  # Gripper Configurations depending on the Object Type , add new force and speed in the Defines if necessary
  # create_gripper_config(gripper_offset=struct(prepick=2, pick=0, place=2), force=0, speed=0, validation=0, object=create_object())
  GRIPPER_CONFIG_MAP.append(create_gripper_config(gripper_offset=struct(prepick=2, pick=0, place=2), force=GRIPPER_FORCE.HALF, speed=GRIPPER_SPEED.MEDIUM, validation=GRIPPER_VALIDATION.ON, object=find_object_by_objectname(Objects.ANY_SAMPLE)))
  GRIPPER_CONFIG_MAP.append(create_gripper_config(gripper_offset=struct(prepick=2, pick=0, place=2), force=GRIPPER_FORCE.FULL, speed=GRIPPER_SPEED.MEDIUM, validation=GRIPPER_VALIDATION.ON, object=find_object_by_objectname(Objects.ANY_RACK)))
  GRIPPER_CONFIG_MAP.append(create_gripper_config(gripper_offset=struct(prepick=2, pick=0, place=2), force=GRIPPER_FORCE.HALF, speed=GRIPPER_SPEED.MEDIUM, validation=GRIPPER_VALIDATION.ON, object=find_object_by_objectname(Objects.CC_SAMPLE)))
  GRIPPER_CONFIG_MAP.append(create_gripper_config(gripper_offset=struct(prepick=3, pick=0, place=3), force=GRIPPER_FORCE.HALF, speed=GRIPPER_SPEED.MEDIUM, validation=GRIPPER_VALIDATION.ON, object=find_object_by_objectname(Objects.HEMA_SAMPLE)))
  GRIPPER_CONFIG_MAP.append(create_gripper_config(gripper_offset=struct(prepick=4, pick=0, place=4), force=GRIPPER_FORCE.HALF, speed=GRIPPER_SPEED.MEDIUM, validation=GRIPPER_VALIDATION.OFF, object=find_object_by_objectname(Objects.TARA_SAMPLE)))
  GRIPPER_CONFIG_MAP.append(create_gripper_config(gripper_offset=struct(prepick=2, pick=0, place=2), force=GRIPPER_FORCE.FULL, speed=GRIPPER_SPEED.MEDIUM, validation=GRIPPER_VALIDATION.ON, object=find_object_by_objectname(Objects.CF_RACK)))
  GRIPPER_CONFIG_MAP.append(create_gripper_config(gripper_offset=struct(prepick=2, pick=0, place=2), force=GRIPPER_FORCE.FULL, speed=GRIPPER_SPEED.MEDIUM, validation=GRIPPER_VALIDATION.ON, object=find_object_by_objectname(Objects.COBAS_RACK)))
  GRIPPER_CONFIG_MAP.append(create_gripper_config(gripper_offset=struct(prepick=0, pick=0, place=0), force=GRIPPER_FORCE.HALF, speed=GRIPPER_SPEED.MEDIUM, validation=GRIPPER_VALIDATION.OFF, object=find_object_by_objectname(Objects.NONE)))
  GRIPPER_CONFIG_MAP.append(create_gripper_config(gripper_offset=struct(prepick=0, pick=0, place=0), force=GRIPPER_FORCE.HALF, speed=GRIPPER_SPEED.MEDIUM, validation=GRIPPER_VALIDATION.OFF, object=find_object_by_objectname(Objects.BUTTON)))
  GRIPPER_CONFIG_MAP.append(create_gripper_config(gripper_offset=struct(prepick=5, pick=25, place=5), force=GRIPPER_FORCE.HALF, speed=GRIPPER_SPEED.MEDIUM, validation=GRIPPER_VALIDATION.OFF, object=find_object_by_objectname(Objects.XN550_DRAWER)))
  # create Patterns like Racks or Magazines
  # easy if you define x and y regarding to the base coordinate system  if not you have to deal with transpose and or invert
  # create_pattern(id=0, pattern_width=[0, 0], pattern_size=[0, 0], blocked=[-1, -1], obj_name=0, direction="X", transpose=False, invert=False, description="default")
  # Objectss: NONE=0, CC_SAMPLE=1, CC_RACK=2, COAG_SAMPLE=3, COAG_RACK=4, HEMA_SAMPLE=5, HEMA_RACK=6, INPUT_RACK=7, CENTRIFUGE_RACK=8, ANY_SAMPLE=9, ANY_RACK=10
  # ITEM_MODEL_MAP.append(create_pattern(id=0, pattern_width=[0, 0], pattern_size=[0, 0], blocked=[-1, -1, -1],  direction="X", transpose=False, invert=False, description="default"))
  # ITEM_MODEL_MAP.append(create_pattern(id=1, pattern_width=[0.06, 0], pattern_size=[3, 1],  direction="X", description="Tara"))
  # ITEM_MODEL_MAP.append(create_pattern(id=2, pattern_width=[0.183, 0.082], pattern_size=[10, 5], description="Sarstedt 50 D17 Rack"))
  # ITEM_MODEL_MAP.append(create_pattern(id=3, pattern_width=[0.153, 0.067], pattern_size=[10, 5], description="Sarstedt 50 D13 Rack"))
  # ITEM_MODEL_MAP.append(create_pattern(id=4, pattern_width=[0.06, 0.06], pattern_size=[3, 3], blocked=[5, -1, -1], description="Hettich Centrifuge Rack"))
  # ITEM_MODEL_MAP.append(create_pattern(id=5, pattern_width=[0.093, 0.093], pattern_size=[2, 2],  description="Hettich Centrifuge Rack Magazin"))
  # ITEM_MODEL_MAP.append(create_pattern(id=6, pattern_width=[0.08, 0.05], pattern_size=[5, 2], description="Sysmex XN 550 Rack"))
  # ITEM_MODEL_MAP.append(create_pattern(id=7, pattern_width=[0.175, 0.078], pattern_size=[8, 4], description="URG Rack 40 D17"))
  # ITEM_MODEL_MAP.append(create_pattern(id=8, pattern_width=[0.092, 0], pattern_size=[5, 1], description="Cobas Rack"))
  # ITEM_MODEL_MAP.append(create_pattern(id=9, pattern_width=[0.245, 0.123], pattern_size=[3, 5], blocked=[9,11,12], description="Cobas Rack Magazin"))
  # ITEM_MODEL_MAP.append(create_pattern(id=10, pattern_width=[0.237, 0.095], pattern_size=[11, 5], description="Atellica Rack 5x11"))
  # ITEM_MODEL_MAP.append(create_pattern(id=11, pattern_width=[0.237, 0.095], pattern_size=[2, 2], description="Sensors LM"))
  # ITEM_MODEL_MAP.append(create_pattern(id=12, pattern_width=[0.18, 0], pattern_size=[10, 1], description="Sysmex CS2500 Rack"))
  # ITEM_MODEL_MAP.append(create_pattern(id=13, pattern_width=[0.310, 0.075], pattern_size=[13, 4], description="URG RACK 52 - Special Input"))
  # ITEM_MODEL_MAP.append(create_pattern(id=14, pattern_width=[0.075, 0.075], pattern_size=[4, 6], description="URG RACK 24 - Special NoK"))
  # ITEM_MODEL_MAP.append(create_pattern(id=15, pattern_width=[0.120, 0], pattern_size=[2, 1], description="XN550 Drawer"))

  ITEM_MODEL_MAP.append(create_pattern(id=0, name="NONE", pattern_width=[0, 0], pattern_size=[0, 0], blocked=[-1, -1, -1],  direction="X", transpose=False, invert=False, description="default"))
  ITEM_MODEL_MAP.append(create_pattern(id=1, name="TARA", pattern_width=[0.06, 0], pattern_size=[3, 1],  direction="X", description="Tara"))
  ITEM_MODEL_MAP.append(create_pattern(id=4, name="CENTRIFUGE", pattern_width=[0.06, 0.06], pattern_size=[3, 3], blocked=[5, -1, -1], description="Hettich Centrifuge Rack"))
  ITEM_MODEL_MAP.append(create_pattern(id=5, name="CENTRIFUGE_MAGAZINE", pattern_width=[0.093, 0.093], pattern_size=[2, 2],  description="Hettich Centrifuge Rack Magazin"))
  ITEM_MODEL_MAP.append(create_pattern(id=6, name="SYSMEX_XN550", pattern_width=[0.08, 0.05], pattern_size=[5, 2], description="Sysmex XN 550 Rack"))
  ITEM_MODEL_MAP.append(create_pattern(id=8, name="COBAS", pattern_width=[0.092, 0], pattern_size=[5, 1], description="Cobas Rack"))
  ITEM_MODEL_MAP.append(create_pattern(id=9, name="COBAS_MAGAZINE", pattern_width=[0.245, 0.123], pattern_size=[3, 5], blocked=[9,11,12], description="Cobas Rack Magazin"))
  ITEM_MODEL_MAP.append(create_pattern(id=13, name="INPUT", pattern_width=[0.310, 0.075], pattern_size=[13, 4], description="URG RACK 52 - Special Input"))
  ITEM_MODEL_MAP.append(create_pattern(id=14, name="NOK", pattern_width=[0.075, 0.075], pattern_size=[4, 6], description="URG RACK 24 - Special NoK"))
  ITEM_MODEL_MAP.append(create_pattern(id=15, name="DRAWER_XN550", pattern_width=[0.120, 0], pattern_size=[2, 1], description="XN550 Drawer"))
  ITEM_MODEL_MAP.append(create_pattern(id=7, name="ARCHIVE", pattern_width=[0.175, 0.078], pattern_size=[8, 4], description="URG Rack 40 D17"))






  # add a "skill" to the robots skillset the control system will send a string with the ls_item and action and here we will look if we have a matching skill to execute
  # the item_modell defines the patterns which have to be used by the robot on multiple racks and or multiple samples in a rackpattern
  # inner pattern is always dependung on the object that has to be moved and the outer pattern is the pattern for the containers where the objects are stored in.
  # if racks have to be handled it is also an inner pattern cause the object to handle is the rack itself
  # create_item(id=0, ls_item="default", frame=p[0,0,0,0,0,0], actionlist=create_action_list([]), item_model=create_item_model(), lm_id=0, description="default")
  # create_item_model(inner=create_pattern(), outer=create_pattern(), description="default")
  # ITEM_MAP.append(create_item(id=1, ls_item="Home", frame=F1_uLM_Home, actionlist=[ActionManipulator.MOVE_TO], description="uLM Move To Home"))
  # ITEM_MAP.append(create_item(id=2, ls_item="InputStation", frame=F2_uLM_Input, actionlist=[ActionManipulator.PICK, ActionManipulator.PLACE], item_model=create_item_model(inner=Patterns.INPUT), description="uLM Pick and Place samples from Input"))
  # ITEM_MAP.append(create_item(id=3, ls_item="InputCapture", frame=F3_Cap_Input, actionlist=[ActionCamera.INSPECT, ActionManipulator.MOVE_TO], description="uLM Inspect samples from Input and Move To Capture Position"))
  # ITEM_MAP.append(create_item(id=4, ls_item="Bin", frame=F4_uLM_Bin, actionlist=[ActionManipulator.PLACE], description="uLM Place Cap to Bin"))
  # ITEM_MAP.append(create_item(id=5, ls_item="StationaryGripper", frame=F5_uLM_Gripper, actionlist=[ActionManipulator.PICK, ActionManipulator.PLACE, ActionManipulator.DECAP, ActionManipulator.MOVE_TO, ActionManipulator.GRASP, ActionManipulator.RELEASE], description=" uLM stationary gripper"))
  # ITEM_MAP.append(create_item(id=6, ls_item="CobasRack", frame=F6_uLM_Cobas_R, actionlist=[ActionManipulator.PICK, ActionManipulator.PLACE], item_model=create_item_model(outer=Patterns.COBAS_MAGAZINE), description="uLM Cobas Racks Pick and Place"))
  # ITEM_MAP.append(create_item(id=7, ls_item="CobasMagazine", frame=F7_uLM_Coba_Mag, actionlist=[ActionManipulator.PICK, ActionManipulator.PLACE], item_model=create_item_model(inner=Patterns.COBAS, outer=Patterns.COBAS_MAGAZINE), description="uLM Cobas Magazine Samples Pick and Place"))
  # ITEM_MAP.append(create_item(id=8, ls_item="DetectCobasRacks", frame=F8_Cap_Cobas_LM, actionlist=[ActionCamera.DETECT_OBJECTS, ActionManipulator.MOVE_TO], lm_id=2, description="uLM Cobas Rack Detection and Move To Capture"))
  # ITEM_MAP.append(create_item(id=9, ls_item="TaraMagazine", frame=F9_uLM_Tara, actionlist=[ActionManipulator.PICK, ActionManipulator.PLACE], item_model=create_item_model(inner=Patterns.TARA), description="uLM Centrifuge Tara Pick and Place"))
  # ITEM_MAP.append(create_item(id=10, ls_item="CentrifugeCapture", frame=F10_Cap_CF, actionlist=[ActionManipulator.MOVE_TO, ActionCamera.DETECT], lm_id=1, description="Centrifuge Device Move to Capture Pos and Detect Landmarks"))
  # ITEM_MAP.append(create_item(id=11, ls_item="Centrifuge", frame=F11_CF_PiPl, actionlist=[ActionManipulator.PICK, ActionManipulator.PLACE], description="Centrifuge Device Rack Pick and Place"))
  # ITEM_MAP.append(create_item(id=12, ls_item="CentrifugeMagazine", frame=F12_uLM_CF_Mag, actionlist=[ActionManipulator.PICK, ActionManipulator.PLACE], item_model=create_item_model(inner=Patterns.CENTRIFUGE, outer=Patterns.CENTRIFUGE_MAGAZINE), description=" uLM Centrifuge Magazin Pick and Place"))
  # ITEM_MAP.append(create_item(id=13, ls_item="CentrifugeRack", frame=F13_uLM_CF_R, actionlist=[ActionManipulator.PICK, ActionManipulator.PLACE], item_model=create_item_model(outer=Patterns.CENTRIFUGE_MAGAZINE), description="uLM Centrifuge Magazin Pick and Place Racks"))
  # ITEM_MAP.append(create_item(id=14, ls_item="DailyArchive", frame=F14_uLM_Archive, actionlist=[ActionManipulator.PICK, ActionManipulator.PLACE], item_model=create_item_model(inner=Patterns.ARCHIVE), description="uLM Pick and Place samples from Archive Rack"))
  # ITEM_MAP.append(create_item(id=15, ls_item="NokRack", frame=F15_uLM_Nok, actionlist=[ActionManipulator.PICK, ActionManipulator.PLACE], item_model=create_item_model(inner=Patterns.NOK), description="uLM Pick and Place samples from Nok Rack"))
  # ITEM_MAP.append(create_item(id=16, ls_item="CobasInput", frame=F16_Cobas_Input, actionlist=[ActionManipulator.PLACE], description="uLM Place Cobasrack in Cobas Device"))
  # ITEM_MAP.append(create_item(id=17, ls_item="CobasInputCapture", frame=F17_Cobas_Cap, actionlist=[ActionCamera.DETECT, ActionManipulator.MOVE_TO], lm_id=3, description="uLM Place Cobasrack in Cobas Device"))
  # ITEM_MAP.append(create_item(id=18, ls_item="XN550Input", frame=F18_XN550_Input, actionlist=[ActionManipulator.PICK, ActionManipulator.PLACE], item_model=create_item_model(inner=Patterns.SYSMEX_XN550, outer=Patterns.DRAWER_XN550), lm_id=4, description="uLM Pick and Place Samples in or out of XN550 Racks"))
  # ITEM_MAP.append(create_item(id=19, ls_item="XN550Capture", frame=F19_XN550_Cap, actionlist=[ActionCamera.DETECT, ActionManipulator.MOVE_TO], lm_id=4, description="uLM Move To and Capture LM XN550"))
  # ITEM_MAP.append(create_item(id=20, ls_item="XN550Drawer", frame=F20_XN550_Draw, actionlist=[ActionManipulator.DRAWER_OPEN, ActionManipulator.DRAWER_CLOSE], item_model=create_item_model(inner=Patterns.DRAWER_XN550), lm_id=4, description="uLM Open and close Drawer XN550"))
  # ITEM_MAP.append(create_item(id=21, ls_item="XN550Button", frame=F21_XN550_Btn, actionlist=[ActionManipulator.PUSH], lm_id=4, description="uLM Push XN550 Button"))
  # ITEM_MAP.append(create_item(id=22, ls_item="AMR", frame=p[0,0,0,0,0,0], actionlist=[ActionAMR.READ, ActionAMR.LOAD_MISSION, ActionAMR.START_MISSION, ActionAMR.NAVIGATE, ActionAMR.ACKNOWLEDGE], description="all AMR actions"))



  # ITEM_MAP.append(create_item(id=31, ls_item="TestLM", frame=TestLM, actionlist=[ActionManipulator.PICK, ActionManipulator.PLACE], item_model=create_item_model(inner=Rack.SYSMEX_CS2500), lm_id=5, description="LM Test"))
  # Fills the Vision Config List with Projectrelated Data
  # workspaceid and skillid are highly robominds related so probably will not stay like this in the future
  # sample detection: dx and dy are used to calculate the positions in a rack and given by the offset which will be applied in order to assign the sample to a place in the rack
  # create_vision_config(workspace_id="", skill_id="", item_id=-1, capture_pos=p[0,0,0,0,0,0], dx=0, dy=0, target_origin=p[0,0,0,0,0,0], selector="default", description="default")
  # VISION_CONFIG_MAP.append(create_vision_config(workspace_id="96017791-f581-4e9e-93da-6951695fccc8", skill_id="8885cfe1-6784-4293-bd26-52ebdc67bf95", capture_pos=F10_Cap_CF, target_origin=p[0,0,0,0,0,0], item_id=11, description="LM Detect CF"))
  # VISION_CONFIG_MAP.append(create_vision_config(workspace_id="96017791-f581-4e9e-93da-6951695fccc8", skill_id="8885cfe1-6784-4293-bd26-52ebdc67bf95", capture_pos=F8_Cap_Cobas_LM, target_origin=p[0,0,0,0,0,0], item_id=8, description="LM Detect Cobas Racks"))
  # VISION_CONFIG_MAP.append(create_vision_config(workspace_id="8f0ad01c-dc36-4fdd-b295-0b6b4a38b89a", skill_id="afdc9e13-ea83-40d6-a805-bb041453d2e5", capture_pos=F3_Cap_Input, target_origin=F2_uLM_Input, item_id=3, description="Lab Solution Input Capture"))
  # VISION_CONFIG_MAP.append(create_vision_config(workspace_id="96017791-f581-4e9e-93da-6951695fccc8", skill_id="8885cfe1-6784-4293-bd26-52ebdc67bf95", capture_pos=F19_XN550_Cap, target_origin=F18_XN550_Input, item_id=18, description="Input XN550"))
  # VISION_CONFIG_MAP.append(create_vision_config(workspace_id="96017791-f581-4e9e-93da-6951695fccc8", skill_id="8885cfe1-6784-4293-bd26-52ebdc67bf95", capture_pos=F19_XN550_Cap, target_origin=POS_Z, item_id=19, description="LM Detect XN550F"))
  # VISION_CONFIG_MAP.append(create_vision_config(workspace_id="96017791-f581-4e9e-93da-6951695fccc8", skill_id="8885cfe1-6784-4293-bd26-52ebdc67bf95", capture_pos=F10_Cap_CF, target_origin=POS_Z, item_id=10, description="LM Detect CF"))
  # VISION_CONFIG_MAP.append(create_vision_config(workspace_id="96017791-f581-4e9e-93da-6951695fccc8", skill_id="8885cfe1-6784-4293-bd26-52ebdc67bf95", capture_pos=F19_XN550_Cap, target_origin=F20_XN550_Draw, item_id=20, description="Drawer XN550"))
  # VISION_CONFIG_MAP.append(create_vision_config(workspace_id="96017791-f581-4e9e-93da-6951695fccc8", skill_id="8885cfe1-6784-4293-bd26-52ebdc67bf95", capture_pos=F19_XN550_Cap, target_origin=F21_XN550_Btn, item_id=21, description="Button XN550"))
  # VISION_CONFIG_MAP.append(create_vision_config(workspace_id="96017791-f581-4e9e-93da-6951695fccc8", skill_id="8885cfe1-6784-4293-bd26-52ebdc67bf95", capture_pos=TestLMCap, target_origin=p[0,0,0,0,0,0], item_id=30, description="Button XN550"))
  # VISION_CONFIG_MAP.append(create_vision_config(workspace_id="96017791-f581-4e9e-93da-6951695fccc8", skill_id="8885cfe1-6784-4293-bd26-52ebdc67bf95", capture_pos=TestLMCap, target_origin=TestLM, item_id=31, description="Button XN550"))

  # VISION_CONFIG_MAP.append(create_vision_config(workspace_id="96017791-f581-4e9e-93da-6951695fccc8", skill_id="8885cfe1-6784-4293-bd26-52ebdc67bf95", target_origin=p[0,0,0,0,0,0], item_id=11, description="LM Detect CF"))
  # VISION_CONFIG_MAP.append(create_vision_config(workspace_id="96017791-f581-4e9e-93da-6951695fccc8", skill_id="8885cfe1-6784-4293-bd26-52ebdc67bf95", target_origin=p[0,0,0,0,0,0], item_id=8, description="LM Detect Cobas Racks"))
  # VISION_CONFIG_MAP.append(create_vision_config(workspace_id="8f0ad01c-dc36-4fdd-b295-0b6b4a38b89a", skill_id="afdc9e13-ea83-40d6-a805-bb041453d2e5", target_origin=F2_uLM_Input, item_id=3, description="Lab Solution Input Capture"))
  # VISION_CONFIG_MAP.append(create_vision_config(workspace_id="96017791-f581-4e9e-93da-6951695fccc8", skill_id="8885cfe1-6784-4293-bd26-52ebdc67bf95", target_origin=F18_XN550_Input, item_id=18, description="Input XN550"))
  # VISION_CONFIG_MAP.append(create_vision_config(workspace_id="96017791-f581-4e9e-93da-6951695fccc8", skill_id="8885cfe1-6784-4293-bd26-52ebdc67bf95", target_origin=POS_Z, item_id=19, description="LM Detect XN550F"))
  # VISION_CONFIG_MAP.append(create_vision_config(workspace_id="96017791-f581-4e9e-93da-6951695fccc8", skill_id="8885cfe1-6784-4293-bd26-52ebdc67bf95", target_origin=POS_Z, item_id=10, description="LM Detect CF"))
  # VISION_CONFIG_MAP.append(create_vision_config(workspace_id="96017791-f581-4e9e-93da-6951695fccc8", skill_id="8885cfe1-6784-4293-bd26-52ebdc67bf95", target_origin=F20_XN550_Draw, item_id=20, description="Drawer XN550"))
  # VISION_CONFIG_MAP.append(create_vision_config(workspace_id="96017791-f581-4e9e-93da-6951695fccc8", skill_id="8885cfe1-6784-4293-bd26-52ebdc67bf95", target_origin=F21_XN550_Btn, item_id=21, description="Button XN550"))
  # VISION_CONFIG_MAP.append(create_vision_config(workspace_id="96017791-f581-4e9e-93da-6951695fccc8", skill_id="8885cfe1-6784-4293-bd26-52ebdc67bf95", target_origin=p[0,0,0,0,0,0], item_id=30, description="Button XN550"))
  # VISION_CONFIG_MAP.append(create_vision_config(workspace_id="96017791-f581-4e9e-93da-6951695fccc8", skill_id="8885cfe1-6784-4293-bd26-52ebdc67bf95", target_origin=TestLM, item_id=31, description="Button XN550"))

  # local inputrack = find_pattern_by_name("INPUT")
  # INSPECT_CONFIG_MAP.append(create_inspect_config(item_id=3, dx=inputrack.pattern_width[0]/(inputrack.pattern_size[0]-1), dy=inputrack.pattern_width[1]/(inputrack.pattern_size[1]-1), rack_size=inputrack.pattern_size , description="Input Capture"))
  # # Fills the Landmark List with Projectrelated Data
  # # create_landmark(lm_id=0, marker_id=-1, marker_size=0.1, marker_type="aruco_7x7", capture_pos=p[0,0,0,0,0,0], init_frame=p[0,0,0,0,0,0], search_offset=[0,0,0], actual_frame=p[0,0,0,0,0,0], description="")
  # LANDMARK_MAP.append(create_landmark(lm_id=1, marker_id=3, marker_size=0.1, marker_type="aruco_7x7", capture_pos = F10_Cap_CF, init_frame=p[-0.617789, -0.065471, 0.07918, 0.020983, -0.012695, 1.512066], search_offset=[0.15, 0.15, 0.1], actual_frame=p[-0.617789, -0.065471, 0.07918, 0.020983, -0.012695, 1.512066], description="LM CF Lid"))
  # LANDMARK_MAP.append(create_landmark(lm_id=2, marker_id=-1, marker_size=0.0085, marker_type="aruco_4x4", capture_pos = F8_Cap_Cobas_LM, init_frame=p[0,0,0,0,0,0], search_offset=[0.15, 0.15, 0.1], actual_frame=POS_Z, description="LM Cobas Rack Detection"))
  # LANDMARK_MAP.append(create_landmark(lm_id=3, marker_id=0, marker_size=0.1, marker_type="aruco_7x7", capture_pos = F17_Cobas_Cap, init_frame=p[-0.667,-0.194,0.100,0,0,0], search_offset=[0.15, 0.15, 0.1], actual_frame=POS_Z, description="LM Cobas Cap"))
  # LANDMARK_MAP.append(create_landmark(lm_id=4, marker_id=4, marker_size=0.1, marker_type="aruco_7x7", capture_pos = F19_XN550_Cap, init_frame=p[0.124,-0.976,0.355,-0.008,0.025,3.131], search_offset=[0.15, 0.15, 0.1], actual_frame=p[0,0,0,0,0,0], description="LM XN550 Cap"))
  # LANDMARK_MAP.append(create_landmark(lm_id=5, marker_id=0, marker_size=0.1, marker_type="aruco_7x7", capture_pos = TestLMCap, init_frame=p[-0.49,-0.144,0.092,0,-0.008,0.001], search_offset=[0.15, 0.15, 0.1], actual_frame=POS_Z, description="LM Test"))
  # # Configuration of all movement related parameters
  # # create_movement(id=0, hh_approach=POS_Z, h_approach=POS_Z, approach=POS_Z, h_target=POS_Z, target=POS_Z, retract=POS_Z, h_retract=POS_Z, hh_retract=POS_Z, h_frame=POS_Z, frame=POS_Z, speed=1, acceleration=1, description="default")
  # MOVEMENT_MAP.append(create_movement(description="TestLMCap", frame=TestLMCap, actionlist=[ActionManipulator.MOVE_TO]))
  # MOVEMENT_MAP.append(create_movement(description="TestLM", frame=TestLM, actionlist=[ActionManipulator.PICK,ActionManipulator.PLACE],
  #         approach=p[0,0,0.1,0,0,0],
  #         retract=p[0,0,0.1,0,0,0]))
  # MOVEMENT_MAP.append(create_movement(description="Home - MOVE_TO", frame=F1_uLM_Home, actionlist=[ActionManipulator.MOVE_TO]))
  # MOVEMENT_MAP.append(create_movement(description="Input - PICK&PLACE", frame=F2_uLM_Input, actionlist=[ActionManipulator.PICK,ActionManipulator.PLACE],
  #         approach=p[0,0,0.1,0,0,0],
  #         retract=p[0,0,0.1,0,0,0]))
  # MOVEMENT_MAP.append(create_movement(description="Capture Input - MOVE_TO", frame=F3_Cap_Input, actionlist=[ActionManipulator.MOVE_TO]))
  # MOVEMENT_MAP.append(create_movement(description="BIN - PLACE", frame=F4_uLM_Bin, actionlist=[ActionManipulator.PLACE],
  #         approach=p[0,0,0.1,0,0,0],
  #         retract=p[0,0,0.1,0,0,0]))
  # MOVEMENT_MAP.append(create_movement(description="Gripper - Move To", frame=F5_uLM_Gripper, actionlist=[ActionManipulator.MOVE_TO],
  #         approach=p[0,0,0.1,0,0,0]))
  # MOVEMENT_MAP.append(create_movement(description="Gripper - Pick", frame=F5_uLM_Gripper, actionlist=[ActionManipulator.PICK],
  #         retract=p[0,0,0.1,0,0,0]))
  # MOVEMENT_MAP.append(create_movement(description="Gripper - Place", frame=F5_uLM_Gripper, actionlist=[ActionManipulator.PLACE],
  #         approach=p[0,0,0.1,0,0,0]))
  # MOVEMENT_MAP.append(create_movement(description="CobasRack Pick & Place", frame=F6_uLM_Cobas_R, actionlist=[ActionManipulator.PICK,ActionManipulator.PLACE],
  #         approach=p[0,0,0.1,0,0,0],
  #         target=p[0,0,0,0,0,d2r(90)],
  #         retract=p[0,0,0.1,0,0,0]))
  # MOVEMENT_MAP.append(create_movement(description="CobasMagazine Pick & Place", frame=F7_uLM_Coba_Mag, actionlist=[ActionManipulator.PICK,ActionManipulator.PLACE],
  #         approach=p[0,0,0.1,0,0,0],
  #         target=p[0,0,0,0,0,-d2r(90)],
  #         retract=p[0,0,0.1,0,0,0]))
  # MOVEMENT_MAP.append(create_movement(description="Capture Position Cobas Landmarks", frame=F8_Cap_Cobas_LM, actionlist=[ActionManipulator.MOVE_TO]))
  # MOVEMENT_MAP.append(create_movement(description="TaraMagazine - PICK & PLACE", frame=F9_uLM_Tara, actionlist=[ActionManipulator.PICK,ActionManipulator.PLACE],
  #         approach=p[0,0,0.13,0,0,0],
  #         target=p[0,0,0,0,0,-d2r(90)],
  #         retract=p[0,0,0.13,0,0,0]))
  # MOVEMENT_MAP.append(create_movement(description="Capture Position - Centrifuge LM", frame=F10_Cap_CF,actionlist=[ActionManipulator.MOVE_TO]))
  # MOVEMENT_MAP.append(create_movement(description="Pick and Place Racks - Centrifuge Lid", frame=F11_CF_PiPl, actionlist=[ActionManipulator.PICK,ActionManipulator.PLACE],
  #         approach=p[0,0,0.3,0,0,0],
  #         retract=p[0,0,0.3,0,0,0]))
  # MOVEMENT_MAP.append(create_movement(description="Pick and Place Samples - Centrifuge on uLM", frame=F12_uLM_CF_Mag, actionlist=[ActionManipulator.PICK,ActionManipulator.PLACE],
  #         approach=p[0,0,0.13,0,0,0],
  #         retract=p[0,0,0.13,0,0,0]
  #         ))
  # MOVEMENT_MAP.append(create_movement(description="Pick and Place Racks - Centrifuge on uLM", frame=F13_uLM_CF_R, actionlist=[ActionManipulator.PICK,ActionManipulator.PLACE],
  #         approach=p[0,0,0.15,0,0,0],
  #         retract=p[0,0,0.15,0,0,0]
  #         ))

  # MOVEMENT_MAP.append(create_movement(description="Pick and Place Samples XN550 Racks in Device", frame=F18_XN550_Input, actionlist=[ActionManipulator.PICK,ActionManipulator.PLACE],
  #         approach=p[0,0,0.1,0,0,0],
  #         target = p[0,0,0,0,0,d2r(90)],
  #         retract=p[0,0,0.1,0,0,0]
  #         ))
  # MOVEMENT_MAP.append(create_movement(description="Capture LM XN550", frame=F19_XN550_Cap, actionlist=[ActionManipulator.MOVE_TO]))
  # MOVEMENT_MAP.append(create_movement(description="Open XN550 Drawer ", frame=F20_XN550_Draw, actionlist=[ActionManipulator.DRAWER_OPEN],
  #         h_approach=p[0.07,0,0.1,0,0,0],
  #         approach=p[0,0,0.1,0,0,0],
  #         target = p[0,0,0,0,0,d2r(90)],
  #         retract=p[0.07,0,0,0,0,0],
  #         h_retract=p[0.07,0,0.1,0,0,0]
  #         ))
  # MOVEMENT_MAP.append(create_movement(description="Close XN550 Drawer ", frame=F20_XN550_Draw, actionlist=[ActionManipulator.DRAWER_CLOSE],
  #         h_approach=p[0.07,0,0.1,0,0,0],
  #         approach=p[0.07,0,0,0,0,0],
  #         target = p[0,0,0,0,0,d2r(90)],
  #         retract=p[0,0,0.1,0,0,0],
  #         h_retract=p[0.07,0,0.1,0,0,0]
  #         ))
  # MOVEMENT_MAP.append(create_movement(description="Push XN550 Button ", frame=F21_XN550_Btn, actionlist=[ActionManipulator.PUSH],
  #         approach=p[0,0,0.15,0,0,0],
  #         retract=p[0,0,0.15,0,0,0]
  #         ))
  # MOVEMENT_MAP.append(create_movement(description="Capture Position 2 Input", frame=F_Cap_Input2,actionlist=[ActionManipulator.MOVE_TO]))



  $ 18 "Script: SCRIPT Objects V0.1.script"
  #*****************************************************
  # customer          :   INTERNAL
  # project name      :
  #****************************************************
  # controller        :   UR
  # software          :   5.17.3
  #****************************************************
  # author            :   P. Koehnke
  # Copyright (c)     :   United Robotics Group
  #                       An der Riede 2
  #                       28816 Stuhr
  #                       Germany
  #****************************************************
  # description       :   object database
  # version:      	:   0.1
  # created           :   09.10.2024
  # updated           :
  #****************************************************
  # modifications     :
  #
  # date              :
  # name              :
  # reason            :
  #****************************************************

  def create_object_2(id=0, name="", type=0, dimension=struct(length=0, width=0, height=0, diameter=0), gripper_offset=p[0,0,0,0,0,0]):
      return struct(id=id, name=name, type=type, dimension=dimension, gripper_offset=gripper_offset)
  end

  OBJ = create_object_2()
  OBJs = make_list(0, create_object_2(), 50)

  OBJs.append(create_object_2(id=1, name="rack centrifuge", type=1, dimension=struct(length=0, width=0, height=0.106, diameter=0.020), gripper_offset=p[0,0,0.095,0,0,2.356]))
  OBJs.append(create_object_2(id=2, name="sample tube 1", type=2, dimension=struct(length=0, width=0, height=0.106, diameter=0.015), gripper_offset=p[0,0,0,0,0,0]))
  OBJs.append(create_object_2(id=3, name="rack sarstedt", type=3, dimension=struct(length=0, width=0, height=0.100, diameter=0.020), gripper_offset=p[0,0,0,0,0,0]))
  OBJs.append(create_object_2(id=4, name="Lab bottle", type=4, dimension=struct(length=0, width=0, height=0.100, diameter=0.030), gripper_offset=p[0,0,0.2,0,0,0]))
  OBJs.append(create_object_2(id=5, name="Vial", type=5, dimension=struct(length=0, width=0, height=0.100, diameter=0.0275), gripper_offset=p[0,0,0,0,0,0]))
  OBJs.append(create_object_2(id=6, name="Container_S", type=6, dimension=struct(length=0.09, width=0.09, height=0.185, diameter=0.080), gripper_offset=p[0,0,0,0,0,0]))
  OBJs.append(create_object_2(id=7, name="Target_container", type=7, dimension=struct(length=0.06, width=0.06, height=0.134, diameter=0.05), gripper_offset=p[0,0,0,0,0,0]))
  OBJs.append(create_object_2(id=8, name="Spatula", type=8, dimension=struct(length=0.03, width=0.03, height=0.23, diameter=0.05), gripper_offset=p[0,0,0,0,0,0]))
  OBJs.append(create_object_2(id=9, name="rack pipet", type=9, dimension=struct(length=0.03, width=0.03, height=0.23, diameter=0.05), gripper_offset=p[0,0,0,0,0,0]))

  def create_jig_2(id=0, name="", type=0, capacity=0, jig_offset=p[0,0,0,0,0,0]):
      # iformation about used jigs
      return struct(id=id, name=name, type=type, capacity=capacity, jig_offset=jig_offset)
  end

  JIG2 = create_jig_2()
  JIGs = make_list(0, create_jig_2(), 20)

  JIGs.append(create_jig_2(id=1, name="3FG", type=1, capacity=1, jig_offset=p[0,0,0,0,0,0]))
  JIGs.append(create_jig_2(id=2, name="jig input", type=2, capacity=1, jig_offset=p[0,0,0,0,0,-3.927]))
  JIGs.append(create_jig_2(id=3, name="jig output", type=3, capacity=1, jig_offset=p[0,0,0,0,0,0.78]))
  JIGs.append(create_jig_2(id=6, name="jig bin", type=6, capacity=1, jig_offset=p[0,0,0,0,0,0]))
  JIGs.append(create_jig_2(id=7, name="jig sarstedt racks", type=7, capacity=1, jig_offset=p[0,0,-0.02,0,0,0]))
  JIGs.append(create_jig_2(id=8, name="NoK Bin", type=8, capacity=1, jig_offset=p[0,0,0,0,0,0]))
  JIGs.append(create_jig_2(id=9, name="Pick bott jig", type=9, capacity=1, jig_offset=p[0,0,0,0,0,0]))
  JIGs.append(create_jig_2(id=10, name="Place bott jig", type=10, capacity=1, jig_offset=p[0,0,0,0,0,0]))
  JIGs.append(create_jig_2(id=11, name="bottle shake jig", type=11, capacity=1, jig_offset=p[0,0,0,0,0,0]))
  JIGs.append(create_jig_2(id=12, name="Pick Vial jig", type=12, capacity=1, jig_offset=p[0,0,0,0,0,0]))
  JIGs.append(create_jig_2(id=13, name="Place Vial jig", type=13, capacity=1, jig_offset=p[0,0,0,0,0,0]))
  JIGs.append(create_jig_2(id=14, name="Liquid transfer jig", type=14, capacity=1, jig_offset=p[0,0,0,0,0,0]))
  JIGs.append(create_jig_2(id=15, name="Pick station jig", type=15, capacity=1, jig_offset=p[0,0,0,0,0,0]))
  JIGs.append(create_jig_2(id=16, name="Place station jig", type=16, capacity=1, jig_offset=p[0,0,0,0,0,0]))
  JIGs.append(create_jig_2(id=17, name="Weigh station jig", type=17, capacity=1, jig_offset=p[0,0,0,0,0,0]))
  JIGs.append(create_jig_2(id=18, name="Pick station 1", type=18, capacity=1, jig_offset=p[0,0,0,0,0,0]))
  JIGs.append(create_jig_2(id=19, name="Pick station 2", type=19, capacity=1, jig_offset=p[0,0,0,0,0,0]))
  JIGs.append(create_jig_2(id=20, name="Pick station 3", type=20, capacity=1, jig_offset=p[0,0,0,0,0,0]))
  JIGs.append(create_jig_2(id=21, name="Tilt station jig", type=21, capacity=1, jig_offset=p[0,0,0,0,0,0]))
  $ 21 "BeforeStarts"
  $ 22 "uLM"
  $ 23 "CMD_Stop≔ False "
  global CMD_Stop=  False
  $ 24 "CMD_Abort≔ False "
  global CMD_Abort=  False
  $ 25 "CMD_Clear≔ False "
  global CMD_Clear=  False
  $ 26 "STATE≔1"
  global STATE=1
  $ 27 "STATE_Info≔''"
  global STATE_Info=""
  $ 28 "ARM_Referenced≔ False "
  global ARM_Referenced=  False
  $ 29 "zero_ftsensor()"
  zero_ftsensor()
  $ 30 "poses init"
  $ 31 "PSE_A≔p[0,0,0,0,0,0]"
  global PSE_A=p[0,0,0,0,0,0]
  $ 32 "PSE_A_H≔p[0,0,0,0,0,0]"
  global PSE_A_H=p[0,0,0,0,0,0]
  $ 33 "PSE_R≔p[0,0,0,0,0,0]"
  global PSE_R=p[0,0,0,0,0,0]
  $ 34 "PSE_R_H≔p[0,0,0,0,0,0]"
  global PSE_R_H=p[0,0,0,0,0,0]
  $ 35 "PSE_T≔p[0,0,0,0,0,0]"
  global PSE_T=p[0,0,0,0,0,0]
  $ 36 "PSE_T_H≔p[0,0,0,0,0,0]"
  global PSE_T_H=p[0,0,0,0,0,0]
  $ 37 "PSE_C_E≔p[0,0,0,0,0,0]"
  global PSE_C_E=p[0,0,0,0,0,0]
  $ 38 "PSE_C_H≔p[0,0,0,0,0,0]"
  global PSE_C_H=p[0,0,0,0,0,0]
  $ 39 "PSE_C_S≔p[0,0,0,0,0,0]"
  global PSE_C_S=p[0,0,0,0,0,0]
  $ 40 "init_home_by_cartesian_pose(p[0,-0.400,0.300,0,0,0])"
  init_home_by_cartesian_pose(p[0,-0.400,0.300,0,0,0])
  $ 41 "Clearing"
  $ 42 "reset_error()"
  reset_error()
  $ 43 "reset_warning()"
  reset_warning()
  $ 44 "uGo"
  $ 46 "ugo_init( True ,'http://192.168.12.120:10001')"
  ugo_init(  True  ,"http://192.168.12.120:10001")
  $ 47 "ugo_update_outputs()"
  ugo_update_outputs()
  $ 48 "App"
  $ 49 "'ADD APPLICATION SPECIFIC COMMANDS'"
  # 'ADD APPLICATION SPECIFIC COMMANDS'
  $ 50 "Tools"
  $ 51 "OBJ_Picked≔gripper_has_object()"
  global OBJ_Picked=gripper_has_object()
  $ 52 "If OBJ_Picked"
  if (OBJ_Picked):
    # begin: URCap Program Node
    #   Source: Robotiq_Grippers, 1.8.4.4844, Robotiq Inc.
    #   Type: Gripper Activate
    $ 53 "Gripper Activate"

    kill rq_gripper_communication_thread
    rq_gripper_communication_thread_started = False

    rq_init_comm_if_connected(9, "1")
    rq_init_comm_if_connected(2, "2")
    rq_init_comm_if_connected(3, "3")
    rq_init_comm_if_connected(4, "4")
    rq_print_connected_grippers()
    rq_gripper_communication_thread = run rq_gripper_communication()

    while(not rq_gripper_communication_thread_started):
        sync()
    end

    rq_set_max_current_for_all_grippers()

    reset_and_activate = False

    rq_activate_all_grippers(False)
    # end: URCap Program Node
  else:
    $ 54 "Else" "noBreak"
    # begin: URCap Program Node
    #   Source: Robotiq_Grippers, 1.8.4.4844, Robotiq Inc.
    #   Type: Gripper Activate
    $ 55 "Gripper Reset and Activate"

    kill rq_gripper_communication_thread
    rq_gripper_communication_thread_started = False

    rq_init_comm_if_connected(9, "1")
    rq_init_comm_if_connected(2, "2")
    rq_init_comm_if_connected(3, "3")
    rq_init_comm_if_connected(4, "4")
    rq_print_connected_grippers()
    rq_gripper_communication_thread = run rq_gripper_communication()

    while(not rq_gripper_communication_thread_started):
        sync()
    end

    rq_set_max_current_for_all_grippers()

    reset_and_activate = True

    rq_activate_all_grippers(True)
    # end: URCap Program Node
  end
  $ 56 "zero_ftsensor()"
  zero_ftsensor()
  $ 57 "EXTT"
  $ 58 "Set GRP_3F_Enable=Off"
  set_standard_digital_out(4, False)
  $ 59 "Set DO[6]=Off"
  set_standard_digital_out(6, False)
  $ 60 "Set GRP_3F_Decap=Off"
  set_standard_digital_out(3, False)
  $ 61 "Set GRP_3F_Cap=Off"
  set_standard_digital_out(2, False)
  $ 62 "Set GRP_3F_Open=Off"
  set_standard_digital_out(5, False)
  $ 63 "PSE_T≔get_tool_free_pose(dir=[0,0,0.150], move_in_base_frame=True)"
  global PSE_T=get_tool_free_pose(dir=[0,0,0.150], move_in_base_frame=True)
  $ 64 "If is_reachable(Base_const, [PSE_T])"
  if (is_reachable(p[0.0,0.0,0.0,0.0,0.0,0.0], [PSE_T])):
    $ 65 "MoveL"
    $ 66 "PSE_T" "breakAfter"
    movel(PSE_T, a=1.2, v=0.15)
  end
  $ 67 "powder dispensing variable init"
  $ 68 "Start_thread≔ False "
  global Start_thread=  False
  $ 69 "vib_mot_thread≔ False "
  global vib_mot_thread=  False
  $ 70 "kp≔0.00005"
  global kp=0.00005
  $ 71 "ki≔0.0005"
  global ki=0.0005
  $ 72 "kd≔0.002"
  global kd=0.002
  $ 73 "dt≔0.02"
  global dt=0.02
  $ 74 "Integral_error≔0"
  global Integral_error=0
  $ 75 "current_error≔0"
  global current_error=0
  $ 76 "previous_error≔0"
  global previous_error=0
  $ 77 "tilt_increment≔0"
  global tilt_increment=0
  $ 79 "diff≔0"
  global diff=0
  $ 80 "current_pose≔get_actual_tcp_pose()"
  global current_pose= get_actual_tcp_pose ()
  $ 81 "Relative_trans≔p[0.4902, -0.65024, -0.22623, 0.019, -0.263, -5.825]"
  global Relative_trans=p[0.4902, -0.65024, -0.22623, 0.019, -0.263, -5.825]
  $ 82 "ContA_plc_offst≔p[-0.00205, 0.02547, 0.03730, -0.03, -2.183, 6.165]"
  global ContA_plc_offst=p[-0.00205, 0.02547, 0.03730, -0.03, -2.183, 6.165]
  $ 83 "PowA_50_offset≔p[0.21808, -0.19943, 0.06584, 0, 0, 0]"
  global PowA_50_offset=p[0.21808, -0.19943, 0.06584, 0, 0, 0]
  while (True):
    $ 84 "Robot Program"
    $ 85 "MAIN"
    $ 86 "command_manager(external_control='uGO', cond_suspend=(ITM_Manipulated and AMR_AtTarget and AMR_Charging and AMR_Battery<40), cond_unsuspend=(AMR_Battery≟60))"
    command_manager(external_control="uGO", cond_suspend=(ITM_Manipulated  and  AMR_AtTarget  and  AMR_Charging  and  AMR_Battery<40), cond_unsuspend=(AMR_Battery == 60))
    $ 87 "log_state(STATE_Info)"
    log_state(STATE_Info)
    $ 88 "Switch STATE"
    switch_1 = STATE
    $ 89 "Case 1"
    if (1 == switch_1):
      $ 90 "Stopping"
      $ 91 "STATE_Info≔'Stopping'"
      global STATE_Info="Stopping"
      $ 92 "end_freedrive_mode()"
      end_freedrive_mode()
      $ 93 "Set"
      set_tcp(p[0.0,0.0,0.161,3.1415,0.0,0.0])
      $ 94 "PSE_T≔get_tool_free_pose(dir=[0,0,0.150], move_in_base_frame=True)"
      global PSE_T=get_tool_free_pose(dir=[0,0,0.150], move_in_base_frame=True)
      $ 95 "If is_reachable(Base_const, [PSE_T])"
      if (is_reachable(p[0.0,0.0,0.0,0.0,0.0,0.0], [PSE_T])):
        $ 96 "MoveL"
        $ 97 "PSE_T" "breakAfter"
        movel(PSE_T, a=1.2, v=0.15)
      end
      $ 98 "do_transition(keep_rxry=OBJ_Picked, r=0)"
      do_transition(keep_rxry=OBJ_Picked, r=0)
      $ 107 "Call Sub_AMR_MiR_V3"
      Sub_AMR_MiR_V3()
      $ 108 "If stopping() and AMR_Done"
      if (stopping()  and  AMR_Done):
        $ 109 "STATE≔2"
        global STATE=2
        $ 110 "ugo_update_outputs()"
        ugo_update_outputs()
      end
    elif (2 == switch_1):
      $ 111 "Case 2"
      $ 112 "Stopped"
      $ 113 "STATE_Info≔'Stopped'"
      global STATE_Info="Stopped"
      $ 114 "Call Sub_AMR_MiR_V3"
      Sub_AMR_MiR_V3()
      $ 115 "If CMD_Reset"
      if (CMD_Reset):
        $ 116 "STATE≔3"
        global STATE=3
        $ 117 "ugo_update_outputs()"
        ugo_update_outputs()
      end
    elif (3 == switch_1):
      $ 118 "Case 3"
      $ 119 " Resetting"
      $ 120 "STATE_Info≔'Resetting'"
      global STATE_Info="Resetting"
      $ 121 "uML"
      $ 122 "reset_error()"
      reset_error()
      $ 123 "reset_warning()"
      reset_warning()
      $ 124 "PROCESS_Step≔0"
      global PROCESS_Step=0
      $ 125 "PROCESS_Info≔''"
      global PROCESS_Info=""
      $ 126 "ARM_Referenced≔ False "
      global ARM_Referenced=  False
      $ 127 "WRK_Done≔ False "
      global WRK_Done=  False
      $ 128 "ITM_Prepared≔ False "
      global ITM_Prepared=  False
      $ 129 "ITM_Manipulated≔ False "
      global ITM_Manipulated=  False
      $ 130 "STP≔0"
      global STP=0
      $ 131 "Action≔0"
      global Action=0
      $ 132 "Action_Info≔''"
      global Action_Info=""
      $ 133 "ITM_ID≔0"
      global ITM_ID=0
      $ 134 "JIG≔0"
      global JIG=0
      $ 135 "JIG_Slot≔0"
      global JIG_Slot=0
      $ 136 "Task_info≔''"
      global Task_info=""
      $ 137 "Set"
      set_tcp(p[0.0,0.0,0.161,3.1415,0.0,0.0])
      $ 138 "App"
      $ 139 "'ADD APPLICATION SPECIFIC COMMANDS'"
      # 'ADD APPLICATION SPECIFIC COMMANDS'
      $ 140 "OBJ_Type≔0"
      global OBJ_Type=0
      $ 141 "OBJ_Nbr≔0"
      global OBJ_Nbr=0
      $ 142 "If CNT_Rack_Output≥50"
      if (CNT_Rack_Output >= 50):
        $ 143 "CNT_Rack_Output≔0"
        global CNT_Rack_Output=0
      end
      $ 144 "TASK≔struct(ID=0, NAVI=struct(target=0, footprint=0, protectiveOff=0, dock=0), WORK=struct(ITM_ID_Src=0, JIG_ID_Src=0, OBJ_Nbr_Src=0, ACT_Src=0, ITM_ID_Tgt=0, JIG_ID_Tgt=0, OBJ_Nbr_Tgt=0, ACT_Tgt=0, OBJ_Type=0))"
      global TASK=struct(ID=0, NAVI=struct(target=0, footprint=0, protectiveOff=0, dock=0), WORK=struct(ITM_ID_Src=0, JIG_ID_Src=0, OBJ_Nbr_Src=0, ACT_Src=0, ITM_ID_Tgt=0, JIG_ID_Tgt=0, OBJ_Nbr_Tgt=0, ACT_Tgt=0, OBJ_Type=0))
      $ 145 "Call Sub_AMR_MiR_V3"
      Sub_AMR_MiR_V3()
      $ 146 "If resetting() and AMR_Done"
      if (resetting()  and  AMR_Done):
        $ 147 "STATE≔4"
        global STATE=4
        $ 148 "ugo_update_outputs()"
        ugo_update_outputs()
      end
    elif (4 == switch_1):
      $ 149 "Case 4"
      $ 150 "Idle"
      $ 151 "STATE_Info≔'Idle'"
      global STATE_Info="Idle"
      $ 152 "If CMD_Start"
      if (CMD_Start):
        $ 153 "STATE≔5"
        global STATE=5
        $ 154 "ugo_update_outputs()"
        ugo_update_outputs()
      end
    elif (5 == switch_1):
      $ 155 "Case 5"
      $ 156 "Starting"
      $ 157 "STATE_Info≔'Starting'"
      global STATE_Info="Starting"
      $ 158 "'ADD COMMANDS WHAT TO START WITH'"
      # 'ADD COMMANDS WHAT TO START WITH'
      $ 159 "Call Sub_AMR_MiR_V3"
      Sub_AMR_MiR_V3()
      $ 160 "get ugo data"
      $ 161 "Assign Tasks"
      $ 162 "TASK.ID = ugo_get_task()"
      TASK.ID = ugo_get_task()
      $ 163 "If TASK.ID≟1"
      if (TASK.ID == 1):
        $ 164 "Task_info≔'Charge'"
        global Task_info="Charge"
        $ 165 "Parameters"
        $ 166 "AMR_PosTarget≔1"
        global AMR_PosTarget=1
      else:
        $ 167 "ElseIf TASK.ID≟9"
        if (TASK.ID == 9):
          $ 168 "'Pick Sarstedt Rack from Variable source'"
          # 'Pick Sarstedt Rack from Variable source'
          $ 169 "Task_info≔'Navigate to Target'"
          global Task_info="Navigate to Target"
          $ 170 "Parameters"
          $ 171 "AMR_PosTarget≔UGO.read_input('00','ITM_ID')"
          global AMR_PosTarget=UGO.read_input("00","ITM_ID")
        else:
          $ 172 "ElseIf TASK.ID≟99"
          if (TASK.ID == 99):
            $ 173 "Task_info≔'Pick rack pipet'"
            global Task_info="Pick rack pipet"
            $ 174 "Parameters"
            $ 175 "ITM_ID≔1"
            global ITM_ID=1
            $ 176 "OBJ_Type≔9"
            global OBJ_Type=9
            $ 177 "JIG≔18"
            global JIG=18
            $ 178 "AMR_PosTarget≔3"
            global AMR_PosTarget=3
          else:
            $ 179 "ElseIf TASK.ID≟98"
            if (TASK.ID == 98):
              $ 180 "Task_info≔'Place rack pipet'"
              global Task_info="Place rack pipet"
              $ 181 "Parameters"
              $ 182 "ITM_ID≔1"
              global ITM_ID=1
              $ 183 "OBJ_Type≔9"
              global OBJ_Type=9
              $ 184 "JIG≔19"
              global JIG=19
              $ 185 "AMR_PosTarget≔2"
              global AMR_PosTarget=2
            else:
              $ 186 "Else" "noBreak"
              $ 187 "set_error(ERROR_WRONG_ORDER)"
              set_error(ERROR_WRONG_ORDER)
            end
          end
        end
      end
      $ 188 "test ugo"
      $ 189 "Wait: 0.2"
      sleep(0.2)
      $ 190 "ugo_update_outputs()"
      ugo_update_outputs()
      $ 191 "If starting() and AMR_Done"
      if (starting()  and  AMR_Done):
        $ 192 "log_message(Task_info, 'New Task: ')"
        log_message(Task_info, "New Task: ")
        $ 193 "log_message(to_str(TASK.ID), 'Task_ID: ')"
        log_message(to_str(TASK.ID), "Task_ID: ")
        $ 194 "do_transition(keep_rxry=OBJ_Picked)"
        do_transition(keep_rxry=OBJ_Picked)
        $ 195 "STATE≔6"
        global STATE=6
        $ 196 "ugo_update_outputs()"
        ugo_update_outputs()
      end
    elif (6 == switch_1):
      $ 197 "Case 6"
      $ 198 "Execute"
      $ 199 "STATE_Info≔'Execute'"
      global STATE_Info="Execute"
      $ 200 "If  not CMD_Hold and not CMD_Suspend"
      global thread_flag_200=0
      thread Thread_if_200():
        $ 201 "Switch PROCESS_Step"
        switch_2 = PROCESS_Step
        $ 202 "Case 0"
        if (0 == switch_2):
          $ 203 "PROCESS_Info≔'process control'"
          global PROCESS_Info="process control"
          $ 204 "log_process(PROCESS_Info)"
          log_process(PROCESS_Info)
          $ 205 "process control"
          $ 206 "If  not AMR_AtTarget"
          if (  not  AMR_AtTarget):
            $ 207 "PROCESS_Step≔1"
            global PROCESS_Step=1
          else:
            $ 208 "ElseIf (( not ITM_Prepared and  not WRK_Done) or (ITM_Prepared and WRK_Done))"
            if (((  not  ITM_Prepared  and    not  WRK_Done)  or  (ITM_Prepared  and  WRK_Done))):
              $ 209 "PROCESS_Step≔2"
              global PROCESS_Step=2
            else:
              $ 210 "ElseIf  not WRK_Done"
              if (  not  WRK_Done):
                $ 211 "PROCESS_Step≔3"
                global PROCESS_Step=3
              else:
                $ 212 "Else" "noBreak"
                $ 213 "task finished"
                $ 214 "PROCESS_Info≔''"
                global PROCESS_Info=""
                $ 215 "STATE≔7"
                global STATE=7
                $ 216 "ugo_update_outputs()"
                ugo_update_outputs()
              end
            end
          end
        elif (1 == switch_2):
          $ 217 "Case 1"
          $ 218 "navigate"
          $ 219 "'MOVING THE uML'"
          # 'MOVING THE uML'
          $ 220 "PROCESS_Info≔'move to target'"
          global PROCESS_Info="move to target"
          $ 221 "log_process(PROCESS_Info)"
          log_process(PROCESS_Info)
          $ 222 "If TASK.ID≟1"
          if (TASK.ID == 1):
            $ 223 "Action≔51"
            global Action=51
          else:
            $ 224 "Else" "noBreak"
            $ 225 "Action≔52"
            global Action=52
          end
          $ 226 "Call Sub_AMR_MiR_V3"
          Sub_AMR_MiR_V3()
          $ 227 "If AMR_Done"
          if (AMR_Done):
            $ 228 "PROCESS_Step≔0"
            global PROCESS_Step=0
          end
        elif (2 == switch_2):
          $ 229 "Case 2"
          $ 230 "prepare"
          $ 231 "'THINGS THAT HAVE TO BE DONE ONCE IN A SEQUENCE,WORKFLOW'"
          # 'THINGS THAT HAVE TO BE DONE ONCE IN A SEQUENCE,WORKFLOW'
          $ 232 "PROCESS_Info≔'prepare for work'"
          global PROCESS_Info="prepare for work"
          $ 233 "log_process(PROCESS_Info)"
          log_process(PROCESS_Info)
          $ 234 "If TASK.WORK.ITM_ID_Src>1"
          if (TASK.WORK.ITM_ID_Src>1):
            $ 235 "ITM_ID≔TASK.WORK.ITM_ID_Src"
            global ITM_ID=TASK.WORK.ITM_ID_Src
          else:
            $ 236 "ElseIf TASK.WORK.ITM_ID_Tgt>1"
            if (TASK.WORK.ITM_ID_Tgt>1):
              $ 237 "ITM_ID≔TASK.WORK.ITM_ID_Tgt"
              global ITM_ID=TASK.WORK.ITM_ID_Tgt
            end
          end
          $ 238 "If  not ARM_Referenced and (ITM_ID≠0)"
          if (  not  ARM_Referenced  and  (ITM_ID != 0)):
            $ 239 "STP≔1"
            global STP=1
          else:
            $ 240 "ElseIf ARM_Referenced or (ITM_ID≟0)"
            if (ARM_Referenced  or  (ITM_ID == 0)):
              $ 241 "STP≔2"
              global STP=2
            end
          end
          $ 242 "Switch STP"
          switch_3 = STP
          $ 243 "Case 1"
          if (1 == switch_3):
            $ 244 "reference"
            $ 245 "STP_Info≔'reference at target position'"
            global STP_Info="reference at target position"
            $ 246 "log_step(STP_Info)"
            log_step(STP_Info)
            $ 247 "If ITM_ID≟1"
            if (ITM_ID == 1):
              $ 248 "CAM_Done≔ True "
              global CAM_Done=  True
            else:
              $ 249 "Else" "noBreak"
              $ 250 "Action≔131"
              global Action=131
              $ 251 "Call Sub_Vision_V18"
              Sub_Vision_V18()
            end
            $ 253 "If CAM_Done and  not ERROR.FLAG"
            if (CAM_Done  and    not  ERROR.FLAG):
              $ 254 "log_step('ARM referenced')"
              log_step("ARM referenced")
              $ 255 "ARM_Referenced≔ True "
              global ARM_Referenced=  True
            end
          elif (2 == switch_3):
            $ 256 "Case 2"
            $ 257 "manipulate"
            $ 258 "STP_Info≔'manipulate item'"
            global STP_Info="manipulate item"
            $ 259 "log_step(STP_Info)"
            log_step(STP_Info)
            $ 260 "'In case pressing button is needed'"
            # 'In case pressing button is needed'
            $ 261 "If found_in_list(ITM_ID, ITM_ID_List)"
            if (found_in_list(ITM_ID, ITM_ID_List)):
              $ 262 "Switch ITM_ID"
              switch_4 = ITM_ID
              $ 263 "Case 0"
              if (0 == switch_4):
                $ 264 "ITM_Manipulated≔ not ITM_Manipulated"
                global ITM_Manipulated=  not  ITM_Manipulated
              elif (1 == switch_4):
                $ 265 "Case 1"
                $ 266 "ITM_Manipulated≔ not ITM_Manipulated"
                global ITM_Manipulated=  not  ITM_Manipulated
              elif (2 == switch_4):
                $ 267 "Case 2"
              else:
                $ 277 "Default Case"
                $ 278 "ITM_Manipulated≔ not ITM_Manipulated"
                global ITM_Manipulated=  not  ITM_Manipulated
              end
            end
          end
          $ 279 "ITM_Prepared≔(ITM_Manipulated or  not found_in_list(ITM_ID, ITM_ID_List)) and (ARM_Referenced or ITM_ID≟0) and  not WRK_Done"
          global ITM_Prepared=(ITM_Manipulated  or    not  found_in_list(ITM_ID, ITM_ID_List))  and  (ARM_Referenced  or  ITM_ID == 0)  and    not  WRK_Done
          $ 280 "STP≔0"
          global STP=0
          $ 281 "STP_Info≔''"
          global STP_Info=""
          $ 282 "PROCESS_Step≔0"
          global PROCESS_Step=0
        elif (3 == switch_2):
          $ 283 "Case 3"
          $ 284 "work"
          $ 285 "'ADD EVERY MACHINE, OBJECT, STATION TO WORK ON'"
          # 'ADD EVERY MACHINE, OBJECT, STATION TO WORK ON'
          $ 286 "Switch ITM_ID"
          switch_3 = ITM_ID
          $ 287 "Case 1"
          if (1 == switch_3):
            $ 288 "uLM"
            $ 289 "If TASK.ID≟12"
            if (TASK.ID == 12):
              $ 290 "fill racks"
              $ 291 "Action≔151"
              global Action=151
              $ 292 "Call Sub_Vision_V18"
              Sub_Vision_V18()
              $ 293 "If  not ERROR.FLAG"
              if (  not  ERROR.FLAG):
                $ 294 "Actions for the task"
                $ 295 "Action≔1"
                global Action=1
                $ 296 "JIG≔2"
                global JIG=2
                $ 297 "JIG_Slot≔CAM_Result[0]"
                global JIG_Slot=CAM_Result[0]
                $ 298 "OBJ_Nbr≔CAM_Result[0]"
                global OBJ_Nbr=CAM_Result[0]
                $ 299 "OBJ_Type≔2"
                global OBJ_Type=2
                $ 300 "Call Sub_Action_V4"
                Sub_Action_V4()
                $ 301 "If OBJ_Picked"
                if (OBJ_Picked):
                  $ 302 "CAM_Result.remove(0)"
                  CAM_Result.remove(0)
                  $ 303 "PRC_TubCounter≔PRC_TubCounter+1"
                  global PRC_TubCounter=PRC_TubCounter+1
                  $ 304 "If PRC_TubCounter%4≟0"
                  if (PRC_TubCounter%4 == 0):
                    $ 305 "JIG_Slot≔4"
                    global JIG_Slot=4
                  else:
                    $ 306 "Else" "noBreak"
                    $ 307 "JIG_Slot≔PRC_TubCounter%4"
                    global JIG_Slot=PRC_TubCounter%4
                  end
                  $ 308 "OBJ_Nbr≔ceil(PRC_TubCounter/4)"
                  global OBJ_Nbr=ceil(PRC_TubCounter/4)
                  $ 309 "Action≔2"
                  global Action=2
                  $ 310 "JIG≔4"
                  global JIG=4
                  $ 311 "Call Sub_Action_V4"
                  Sub_Action_V4()
                  $ 312 "Action≔151"
                  global Action=151
                  $ 313 "Call Sub_Vision_V18"
                  Sub_Vision_V18()
                end
              end
              $ 314 "If (CAM_Captures≥CAM_PRM_Retries) or (PRC_TubCounter≥32)"
              if ((CAM_Captures >= CAM_PRM_Retries)  or  (PRC_TubCounter >= 32)):
                $ 315 "PROCESS_Step≔0"
                global PROCESS_Step=0
                $ 316 "WRK_Done≔ True "
                global WRK_Done=  True
              end
            else:
              $ 317 "ElseIf TASK.ID≟49"
              if (TASK.ID == 49):
                $ 318 "Pick Powder container"
                $ 319 "Action≔131"
                global Action=131
                $ 320 "Call Sub_Vision_V18"
                Sub_Vision_V18()
                $ 321 "Action≔35"
                global Action=35
                $ 322 "Call Sub_Action_V4"
                Sub_Action_V4()
                $ 323 "PROCESS_Step≔0"
                global PROCESS_Step=0
                $ 324 "WRK_Done≔ True "
                global WRK_Done=  True
              else:
                $ 325 "ElseIf TASK.ID≟50"
                if (TASK.ID == 50):
                  $ 326 "Decap containers"
                  $ 327 "Action≔36"
                  global Action=36
                  $ 328 "Call Sub_Action_V4"
                  Sub_Action_V4()
                  $ 329 "PROCESS_Step≔0"
                  global PROCESS_Step=0
                  $ 330 "WRK_Done≔ True "
                  global WRK_Done=  True
                else:
                  $ 331 "ElseIf TASK.ID≟51"
                  if (TASK.ID == 51):
                    $ 332 "Detect Spatula and transfer powder"
                    $ 333 "Action≔131"
                    global Action=131
                    $ 334 "Call Sub_Vision_V18"
                    Sub_Vision_V18()
                    $ 335 "Action≔37"
                    global Action=37
                    $ 336 "Call Sub_Action_V4"
                    Sub_Action_V4()
                    $ 337 "PROCESS_Step≔0"
                    global PROCESS_Step=0
                    $ 338 "WRK_Done≔ True "
                    global WRK_Done=  True
                  else:
                    $ 339 "ElseIf TASK.ID≟52"
                    if (TASK.ID == 52):
                      $ 340 "Pick PowderA container"
                      $ 341 "Action≔131"
                      global Action=131
                      $ 342 "Call Sub_Vision_V18"
                      Sub_Vision_V18()
                      $ 343 "Action≔38"
                      global Action=38
                      $ 344 "Call Sub_Action_V4"
                      Sub_Action_V4()
                      $ 345 "PROCESS_Step≔0"
                      global PROCESS_Step=0
                      $ 346 "WRK_Done≔ True "
                      global WRK_Done=  True
                    else:
                      $ 347 "ElseIf TASK.ID≟53"
                      if (TASK.ID == 53):
                        $ 348 "Decap containerA"
                        $ 349 "Action≔39"
                        global Action=39
                        $ 350 "Call Sub_Action_V4"
                        Sub_Action_V4()
                        $ 351 "PROCESS_Step≔0"
                        global PROCESS_Step=0
                        $ 352 "WRK_Done≔ True "
                        global WRK_Done=  True
                      else:
                        $ 353 "ElseIf TASK.ID≟54"
                        if (TASK.ID == 54):
                          $ 354 "Dispense PowderA"
                          $ 355 "Action≔131"
                          global Action=131
                          $ 356 "Call Sub_Vision_V18"
                          Sub_Vision_V18()
                          $ 357 "Action≔40"
                          global Action=40
                          $ 358 "Call Sub_Action_V4"
                          Sub_Action_V4()
                          $ 359 "PROCESS_Step≔0"
                          global PROCESS_Step=0
                          $ 360 "WRK_Done≔ True "
                          global WRK_Done=  True
                        else:
                          $ 361 "ElseIf TASK.ID≟54"
                          if (TASK.ID == 54):
                            $ 362 "Dispense PowderA"
                            $ 363 "Action≔131"
                            global Action=131
                            $ 364 "Call Sub_Vision_V18"
                            Sub_Vision_V18()
                            $ 365 "Action≔40"
                            global Action=40
                            $ 366 "Call Sub_Action_V4"
                            Sub_Action_V4()
                            $ 367 "PROCESS_Step≔0"
                            global PROCESS_Step=0
                            $ 368 "WRK_Done≔ True "
                            global WRK_Done=  True
                          else:
                            $ 369 "ElseIf TASK.ID≟99"
                            if (TASK.ID == 99):
                              $ 370 "Pick rack pipet"
                              $ 371 "Action≔131"
                              global Action=131
                              $ 372 "Call Sub_Vision_V18"
                              Sub_Vision_V18()
                              $ 373 "Action≔5"
                              global Action=5
                              $ 374 "Call Sub_Action_V4"
                              Sub_Action_V4()
                              $ 375 "PROCESS_Step≔0"
                              global PROCESS_Step=0
                              $ 376 "WRK_Done≔ True "
                              global WRK_Done=  True
                            else:
                              $ 377 "ElseIf TASK.ID≟98"
                              if (TASK.ID == 98):
                                $ 378 "Pick rack pipet"
                                $ 379 "Action≔131"
                                global Action=131
                                $ 380 "Call Sub_Vision_V18"
                                Sub_Vision_V18()
                                $ 381 "Action≔6"
                                global Action=6
                                $ 382 "Call Sub_Action_V4"
                                Sub_Action_V4()
                                $ 383 "PROCESS_Step≔0"
                                global PROCESS_Step=0
                                $ 384 "WRK_Done≔ True "
                                global WRK_Done=  True
                              end
                            end
                          end
                        end
                      end
                    end
                  end
                end
              end
            end
          elif (2 == switch_3):
            $ 385 "Case 2"
          elif (5 == switch_3):
            $ 427 "Case 5"
          elif (20 == switch_3):
            $ 435 "Case 20"
          elif (43 == switch_3):
            $ 497 "Case 43"
          else:
            $ 505 "Default Case"
            $ 506 "WRK_Done≔ True "
            global WRK_Done=  True
            $ 507 "PROCESS_Step≔0"
            global PROCESS_Step=0
          end
        end
        thread_flag_200 = 1
      end
      if (  not  CMD_Hold and not CMD_Suspend):
        global thread_handler_200=run Thread_if_200()
        while (thread_flag_200 == 0):
          if not(  not  CMD_Hold and not CMD_Suspend):
            kill thread_handler_200
            thread_flag_200 = 2
          else:
            sync()
          end
        end
      else:
        thread_flag_200 = 2
      end
      $ 508 "If CMD_Hold"
      if (CMD_Hold):
        $ 509 "STATE≔9"
        global STATE=9
        $ 510 "ugo_update_outputs()"
        ugo_update_outputs()
      else:
        $ 511 "ElseIf CMD_Suspend"
        if (CMD_Suspend):
          $ 512 "STATE≔12"
          global STATE=12
          $ 513 "ugo_update_outputs()"
          ugo_update_outputs()
        end
      end
    elif (7 == switch_1):
      $ 514 "Case 7"
      $ 515 "Completing"
      $ 516 "STATE_Info≔'Completing'"
      global STATE_Info="Completing"
      $ 517 "'ADD COMMANDS FOR COMPLETING THE PROCESS'"
      # 'ADD COMMANDS FOR COMPLETING THE PROCESS'
      $ 518 "do_transition(keep_rxry=OBJ_Picked)"
      do_transition(keep_rxry=OBJ_Picked)
      $ 519 "Call Sub_AMR_MiR_V3"
      Sub_AMR_MiR_V3()
      $ 520 "If completing() and AMR_Done"
      if (completing()  and  AMR_Done):
        $ 521 "STATE≔8"
        global STATE=8
        $ 522 "ugo_update_outputs()"
        ugo_update_outputs()
      end
    elif (8 == switch_1):
      $ 523 "Case 8"
      $ 524 "Complete"
      $ 525 "STATE_Info≔'Complete'"
      global STATE_Info="Complete"
      $ 526 "If CMD_Reset"
      if (CMD_Reset):
        $ 527 "STATE≔3"
        global STATE=3
        $ 528 "ugo_update_outputs()"
        ugo_update_outputs()
      end
    elif (9 == switch_1):
      $ 529 "Case 9"
      $ 530 "Holding"
      $ 531 "STATE_Info≔'Holding'"
      global STATE_Info="Holding"
      $ 532 "stopl(0.5)"
      stopl(0.5)
      $ 533 "Call Sub_AMR_MiR_V3"
      Sub_AMR_MiR_V3()
      $ 534 "If holding() and AMR_Done"
      if (holding()  and  AMR_Done):
        $ 535 "STATE≔10"
        global STATE=10
        $ 536 "ugo_update_outputs()"
        ugo_update_outputs()
      end
    elif (10 == switch_1):
      $ 537 "Case 10"
      $ 538 "Held"
      $ 539 "STATE_Info≔'Held'"
      global STATE_Info="Held"
      $ 540 "If CMD_Unhold"
      if (CMD_Unhold):
        $ 541 "end_freedrive_mode()"
        end_freedrive_mode()
        $ 542 "STATE≔11"
        global STATE=11
        $ 543 "ugo_update_outputs()"
        ugo_update_outputs()
      else:
        $ 544 "ElseIf FNC_Freedrive"
        if (FNC_Freedrive):
          $ 545 "freedrive_mode()"
          freedrive_mode()
        else:
          $ 546 "Else" "noBreak"
          $ 547 "end_freedrive_mode()"
          end_freedrive_mode()
        end
      end
    elif (11 == switch_1):
      $ 548 "Case 11"
      $ 549 "Unholding"
      $ 550 "STATE_Info≔'Unholding'"
      global STATE_Info="Unholding"
      $ 551 "Clearing"
      $ 552 "Switch ERROR.ID"
      switch_2 = ERROR.ID
      $ 553 "Case 1002"
      if (1002 == switch_2):
        $ 554 "AMR_AtTarget≔ False "
        global AMR_AtTarget=  False
        $ 555 "ARM_Referenced≔ False "
        global ARM_Referenced=  False
        $ 556 "ITM_Prepared≔ False "
        global ITM_Prepared=  False
        $ 557 "PROCESS_Step≔1"
        global PROCESS_Step=1
      elif (2007 == switch_2):
        $ 558 "Case 2007"
        $ 559 "PROCESS_Step≔1"
        global PROCESS_Step=1
      end
      $ 560 "reset_error()"
      reset_error()
      $ 561 "reset_warning()"
      reset_warning()
      $ 562 "OBJ_Picked≔gripper_has_object()"
      global OBJ_Picked=gripper_has_object()
      $ 563 "Call Sub_AMR_MiR_V3"
      Sub_AMR_MiR_V3()
      $ 564 "If unholding() and AMR_Done"
      if (unholding()  and  AMR_Done):
        $ 565 "STATE≔6"
        global STATE=6
        $ 566 "ugo_update_outputs()"
        ugo_update_outputs()
      end
    elif (12 == switch_1):
      $ 567 "Case 12"
      $ 568 "Suspending"
      $ 569 "STATE_Info≔'Suspending'"
      global STATE_Info="Suspending"
      $ 570 "PROCESS_Info≔str_cat(PROCESS_Info, ' suspended')"
      global PROCESS_Info=str_cat(PROCESS_Info, " suspended")
      $ 571 "If suspending()"
      if (suspending()):
        $ 572 "STATE≔13"
        global STATE=13
        $ 573 "ugo_update_outputs()"
        ugo_update_outputs()
      end
    elif (13 == switch_1):
      $ 574 "Case 13"
      $ 575 "Suspended"
      $ 576 "STATE_Info≔'Suspended'"
      global STATE_Info="Suspended"
      $ 577 "Call Sub_AMR_MiR_V3"
      Sub_AMR_MiR_V3()
      $ 578 "If CMD_Unsuspend"
      if (CMD_Unsuspend):
        $ 579 "STATE≔14"
        global STATE=14
        $ 580 "ugo_update_outputs()"
        ugo_update_outputs()
      end
    elif (14 == switch_1):
      $ 581 "Case 14"
      $ 582 "Unsuspending"
      $ 583 "STATE_Info≔'Unsuspending'"
      global STATE_Info="Unsuspending"
      $ 584 "PROCESS_Step≔0"
      global PROCESS_Step=0
      $ 585 "If unsuspending()"
      if (unsuspending()):
        $ 586 "STATE≔6"
        global STATE=6
        $ 587 "ugo_update_outputs()"
        ugo_update_outputs()
      end
    elif (15 == switch_1):
      $ 588 "Case 15"
      $ 589 "Aborting"
      $ 590 "STATE_Info≔'Aborting'"
      global STATE_Info="Aborting"
      $ 591 "If aborting()"
      if (aborting()):
        $ 592 "STATE≔16"
        global STATE=16
        $ 593 "ugo_update_outputs()"
        ugo_update_outputs()
      end
    elif (16 == switch_1):
      $ 594 "Case 16"
      $ 595 "Aborted"
      $ 596 "STATE_Info≔'Aborted'"
      global STATE_Info="Aborted"
      $ 597 "If CMD_Clear"
      if (CMD_Clear):
        $ 598 "STATE≔17"
        global STATE=17
        $ 599 "ugo_update_outputs()"
        ugo_update_outputs()
      end
    elif (17 == switch_1):
      $ 600 "Case 17"
      $ 601 "Clearing"
      $ 602 "STATE_Info≔'Clearing'"
      global STATE_Info="Clearing"
      $ 603 "Clearing"
      $ 604 "reset_warning()"
      reset_warning()
      $ 605 "reset_error()"
      reset_error()
      $ 606 "If clearing()"
      if (clearing()):
        $ 607 "STATE≔2"
        global STATE=2
        $ 608 "ugo_update_outputs()"
        ugo_update_outputs()
      end
    end
    $ 609 "log_state(STATE_Info)"
    log_state(STATE_Info)
    $ 610 "log_warning(WARNING.MSG)"
    log_warning(WARNING.MSG)
    $ 611 "log_error(ERROR.MSG)"
    log_error(ERROR.MSG)
    $ 612 "Times"
    $ 613 "Switch STATE"
    switch_1 = STATE
    $ 614 "Case 1"
    if (1 == switch_1):
      $ 615 "TM_St_Stopping≔get_time(STATE_Times[STATE-1])"
      global TM_St_Stopping=get_time(STATE_Times[STATE-1])
    elif (2 == switch_1):
      $ 616 "Case 2"
      $ 617 "TM_St_Stopped≔get_time(STATE_Times[STATE-1])"
      global TM_St_Stopped=get_time(STATE_Times[STATE-1])
    elif (3 == switch_1):
      $ 618 "Case 3"
      $ 619 "TM_St_Resetting≔get_time(STATE_Times[STATE-1])"
      global TM_St_Resetting=get_time(STATE_Times[STATE-1])
    elif (4 == switch_1):
      $ 620 "Case 4"
      $ 621 "TM_St_Idle≔get_time(STATE_Times[STATE-1])"
      global TM_St_Idle=get_time(STATE_Times[STATE-1])
    elif (5 == switch_1):
      $ 622 "Case 5"
      $ 623 "TM_St_Starting≔get_time(STATE_Times[STATE-1])"
      global TM_St_Starting=get_time(STATE_Times[STATE-1])
    elif (6 == switch_1):
      $ 624 "Case 6"
      $ 625 "TM_St_Execute≔get_time(STATE_Times[STATE-1])"
      global TM_St_Execute=get_time(STATE_Times[STATE-1])
    elif (7 == switch_1):
      $ 626 "Case 7"
      $ 627 "TM_St_Completin≔get_time(STATE_Times[STATE-1])"
      global TM_St_Completin=get_time(STATE_Times[STATE-1])
    elif (8 == switch_1):
      $ 628 "Case 8"
      $ 629 "TM_St_Complete≔get_time(STATE_Times[STATE-1])"
      global TM_St_Complete=get_time(STATE_Times[STATE-1])
    elif (9 == switch_1):
      $ 630 "Case 9"
      $ 631 "TM_St_Holding≔get_time(STATE_Times[STATE-1])"
      global TM_St_Holding=get_time(STATE_Times[STATE-1])
    elif (10 == switch_1):
      $ 632 "Case 10"
      $ 633 "TM_St_Held≔get_time(STATE_Times[STATE-1])"
      global TM_St_Held=get_time(STATE_Times[STATE-1])
    elif (11 == switch_1):
      $ 634 "Case 11"
      $ 635 "TM_St_Unholding≔get_time(STATE_Times[STATE-1])"
      global TM_St_Unholding=get_time(STATE_Times[STATE-1])
    elif (12 == switch_1):
      $ 636 "Case 12"
      $ 637 "TM_St_Suspendin≔get_time(STATE_Times[STATE-1])"
      global TM_St_Suspendin=get_time(STATE_Times[STATE-1])
    elif (13 == switch_1):
      $ 638 "Case 13"
      $ 639 "TM_St_Suspended≔get_time(STATE_Times[STATE-1])"
      global TM_St_Suspended=get_time(STATE_Times[STATE-1])
    elif (14 == switch_1):
      $ 640 "Case 14"
      $ 641 "TM_St_Unsuspend≔get_time(STATE_Times[STATE-1])"
      global TM_St_Unsuspend=get_time(STATE_Times[STATE-1])
    elif (15 == switch_1):
      $ 642 "Case 15"
      $ 643 "TM_St_Aborting≔get_time(STATE_Times[STATE-1])"
      global TM_St_Aborting=get_time(STATE_Times[STATE-1])
    elif (16 == switch_1):
      $ 644 "Case 16"
      $ 645 "TM_St_Aborted≔get_time(STATE_Times[STATE-1])"
      global TM_St_Aborted=get_time(STATE_Times[STATE-1])
    elif (17 == switch_1):
      $ 646 "Case 17"
      $ 647 "TM_St_Clearing≔get_time(STATE_Times[STATE-1])"
      global TM_St_Clearing=get_time(STATE_Times[STATE-1])
    end
    $ 649 "Wait: 0.1"
    sleep(0.1)
  end
end
